(* Logix 5000 project; controller NWGG 1756-L72 rev 35.12; software revision 35.00 *)

TASK _2_MAIN (event, rate 10 ms, priority 15, watchdog 500 ms) : _2_MAIN
TASK Development (event, rate 10 ms, priority 10, watchdog 500 ms) : Main
TASK MainTask (continuous, watchdog 500 ms) : MainProgram
TASK SeedCleaning (event, rate 10 ms, priority 10, watchdog 500 ms) : Amp_Guages
TASK SeedLoadout (event, rate 10 ms, priority 10, watchdog 500 ms) : SeedLoadoutMain, Scale
TASK Test (event, rate 10 ms, priority 10, watchdog 500 ms) : Test
TASK UpdateBinConfig (event, rate 10 ms, priority 10, watchdog 500 ms)

MODULES
   Local : 1756-L72 (ICP 3, rev 35.12)
      R0S3_IA16 : 1756-IA16 (ICP 0, rev 3.1, Input RPI 20 ms)
      R0S2_IA16 : 1756-IA16 (ICP 1, rev 3.1, Input RPI 20 ms)
      R0S5_OA16I : 1756-OA16I (ICP 5, rev 3.1, Output RPI 20 ms)
      R0S6_OA16I : 1756-OA16I (ICP 6, rev 3.1, Output RPI 20 ms)
      R0S1_EN2TR : vendor 1 type 12 code 200 (ICP 4, Ethernet 192.10.21.33, rev 5.1)
         Treater_PLC : vendor 1 type 14 code 107 (Ethernet 192.10.21.15, rev 28.12, $43c9857a$ RPI 20 ms)
         LCP101_ETAP : 1783-ETAP (Ethernet 192.10.21.22, rev 2.1)
         Concrete_PLC : 1769-L35E Ethernet Port (Ethernet 192.10.21.32, rev 18.1)
            Concrete_PLC_Controller : vendor 1 type 14 code 65 (CompactLogixL35Controller 0, rev 18.1, $0a5c8464$ RPI 20 ms, $a6a510d7$ RPI 20 ms, $5be82f5e$ RPI 20 ms, $3e907429$ RPI 20 ms, $784e80a8$ RPI 20 ms, $ecd2168b$ RPI 100 ms, $00c6bec2$ RPI 20 ms, $fbd2347d$ RPI 20 ms, $adf8042c$ RPI 20 ms)
         Cimbria_Fan : PowerFlex 525-EENET (Ethernet 192.10.21.43, rev 4.1, Output RPI 20 ms)
         LCP103_4 : 1794-AENTR (Ethernet 192.10.21.39, rev 1.1, Output RPI 20 ms)
             : 1794-IA16 (Flex 2, rev 1.1)
            INPUT3 : 1794-IB16 (Flex 3, rev 1.1)
            CT_INPUT : 1794-IE12 (Flex 0, rev 1.1, Output RPI 80 ms)
            CT_INPUT2 : 1794-IE12 (Flex 1, rev 1.1, Output RPI 80 ms)
         R5M4_AENTR : 1794-AENTR (Ethernet 192.10.21.25, rev 1.1, Output RPI 20 ms)
            R5S3_IE8 : vendor 1 type 10 code 25 (Flex 3, rev 2.1, Input RPI 80 ms)
            R5S1_OE4 : 1794-OE4 (Flex 1, rev 2.1, Output RPI 80 ms)
            R5S0_OE4 : 1794-OE4 (Flex 0, rev 2.1, Output RPI 80 ms)
            R5S2_IE8 : vendor 1 type 10 code 25 (Flex 2, rev 2.1, Input RPI 80 ms)
         R4M2_AENTR : 1794-AENTR (Ethernet 192.10.21.27, rev 1.1, Output RPI 20 ms)
            R4S3_IA16 : 1794-IA16 (Flex 3, rev 1.1)
            R4S4_IA16 : 1794-IA16 (Flex 4, rev 1.1)
            R4SO_IA16 : 1794-IA16 (Flex 0, rev 1.1)
            R4S2_IA16 : 1794-IA16 (Flex 2, rev 1.1)
            R4S1_IA16 : 1794-IA16 (Flex 1, rev 1.1)
         DISTRIBUTION : 1794-AENTR (Ethernet 192.10.21.28, rev 1.1, Output RPI 20 ms)
            R5S1_OW8 : 1794-OW8 (Flex 1, rev 1.1)
            R5S0 : 1794-IA16 (Flex 0, rev 1.1)
         R4M3_AENTR : 1794-AENTR (Ethernet 192.10.21.26, rev 1.1, Output RPI 20 ms)
            R4S1_OA16 : vendor 1 type 7 code 48 (Flex 1, rev 1.1)
            R4S4_OA16 : vendor 1 type 7 code 48 (Flex 4, rev 1.1)
            R4S0_OA16 : vendor 1 type 7 code 48 (Flex 0, rev 1.1)
            R4S2_OA16 : vendor 1 type 7 code 48 (Flex 2, rev 1.1)
            R4S3_OA16 : vendor 1 type 7 code 48 (Flex 3, rev 1.1)
         R3M1_AENTR : 1794-AENTR (Ethernet 192.10.21.24, rev 1.1, Output RPI 20 ms)
            R3S1_OA16 : vendor 1 type 7 code 48 (Flex 1, rev 1.1)
            R3S3_OA16 : vendor 1 type 7 code 48 (Flex 3, rev 1.1)
            R3S0_IA16 : 1794-IA16 (Flex 0, rev 1.1)
            R3S2_IA16 : 1794-IA16 (Flex 2, rev 1.1)
         Stratix_5700 : vendor 1 type 12 code 241 (Ethernet 192.10.21.200, rev 4.1, Output RPI 1000 ms)
         AveryWT_Bay1 : ETHERNET-MODULE (Ethernet 192.10.21.70, rev 1.1, Output RPI 10 ms)
         AveryWT_Bay2 : ETHERNET-MODULE (Ethernet 192.10.21.71, rev 1.1, Output RPI 10 ms)
         R2S0_AENTR : vendor 1 type 12 code 228 (Ethernet 192.10.21.21, rev 1.1)
            R2S3_NI8 : vendor 1 type 117 code 6 (SLCChassis 3, rev 1.1, StandardDataDriven RPI 20 ms)
            R2S1_OA16 : vendor 1 type 116 code 24 (SLCChassis 1, rev 1.1, StandardDataDriven RPI 20 ms)
            R2S4_NI8 : vendor 1 type 117 code 6 (SLCChassis 4, rev 1.1, StandardDataDriven RPI 20 ms)
            R2S5_NI8 : vendor 1 type 117 code 6 (SLCChassis 5, rev 1.1, StandardDataDriven RPI 20 ms)
         R1S0_AENTR : vendor 1 type 12 code 228 (Ethernet 192.10.21.20, rev 1.1)
            R1S5_IA16 : vendor 1 type 116 code 3 (SLCChassis 5, rev 1.1, StandardDataDriven RPI 20 ms)
            R1S9_OA161 : vendor 1 type 116 code 24 (SLCChassis 10, rev 1.1, StandardDataDriven RPI 20 ms)
            R1S2_IA16 : vendor 1 type 116 code 3 (SLCChassis 2, rev 1.1, StandardDataDriven RPI 20 ms)
            R1S6_IA16 : vendor 1 type 116 code 3 (SLCChassis 6, rev 1.1, StandardDataDriven RPI 20 ms)
            R1S4_IA16 : vendor 1 type 116 code 3 (SLCChassis 4, rev 1.1, StandardDataDriven RPI 20 ms)
            R1S7_IA16 : vendor 1 type 116 code 3 (SLCChassis 7, rev 1.1, StandardDataDriven RPI 20 ms)
            R1S9_OA163 : vendor 1 type 116 code 24 (SLCChassis 12, rev 1.1, StandardDataDriven RPI 20 ms)
            R1S1_IA16 : vendor 1 type 116 code 3 (SLCChassis 1, rev 1.1, StandardDataDriven RPI 20 ms)
            R1S8_IA16 : vendor 1 type 116 code 3 (SLCChassis 8, rev 1.1, StandardDataDriven RPI 20 ms)
            R1S9_OA162 : vendor 1 type 116 code 24 (SLCChassis 11, rev 1.1, StandardDataDriven RPI 20 ms)
            R1S9_OA16 : vendor 1 type 116 code 24 (SLCChassis 9, rev 1.1, StandardDataDriven RPI 20 ms)
            R1S3_IA16 : vendor 1 type 116 code 3 (SLCChassis 3, rev 1.1, StandardDataDriven RPI 20 ms)
      Analog_Input : 1756-IF8 (ICP 2, rev 1.1, Input RPI 100 ms)
END_MODULES

TYPE udt_Andco_Remote_Out :
STRUCT
   Close : BOOL;
   Open : BOOL;
END_STRUCT
END_TYPE

TYPE udt_Andco_Values :
STRUCT
   Faulted : BOOL;
   Closed : BOOL;
   Values_Updated : BOOL;
   Fully_Open : BOOL;
   Com_Fault : BOOL;
   Open_Gate : BOOL;
   Close_Gate : BOOL;
   Cal_Gate : BOOL;
   Move_Gate : BOOL;
   Cal_Status : DINT;
   Raw_Position : DINT;
   Max_Position : DINT;
   Preact : DINT;
   Tolerance : DINT;
   Percent_Open : REAL;
   New_Pos : INT;
   Width : REAL;
   Rate : REAL;
   Pounds_Per_Inch : REAL;
   New_Rate : REAL;
   Set_New_Rate : BOOL;
   Display_New_Rate_Screen : BOOL;
   Analog : BOOL;
   Min_Position : DINT;
   Length : REAL;
   InchesOpen : REAL;
   AnalogValue : DINT;
END_STRUCT
END_TYPE

TYPE udt_Bin_Rate_Cal_Points :
STRUCT
   Andco_Position : INT;
   Rate : INT;
END_STRUCT
END_TYPE

TYPE udt_Clean_Seed_Bin :
STRUCT
   In_Use : BOOL;
   Bin_Name : STRING;
   Andco : udt_Andco_Values;
   Required_Clean_Belt : DINT;
   Required_Treat_Belt : DINT;
   Required_Transfer_Belt : DINT;
   Clean_Legs_Rqd : DINT;
   K_Valves_On_Treat : DINT;
   K_Valves_On_Clean : DINT;
   Concrete_Bin : BOOL;
   High_Bindicator : BOOL;
   Low_Bindicator : BOOL;
   Use_For_Clean : BOOL;
   Use_For_Treated : BOOL;
   Use_For_Transfer : BOOL;
   Cal_Mode : BOOL;
   Time_To_Treater : REAL;
   Time_To_Clean : REAL;
   Auger : BOOL;
   Current_Product : STRING;
   Capacity : DINT;
   Current_Amount : DINT;
END_STRUCT
END_TYPE

TYPE udt_Color :
STRUCT
   Color : INT;
   Duration : INT;
END_STRUCT
END_TYPE

TYPE udt_Cyclone :
STRUCT
   Start_Both_Fans : BOOL;
   Start_Cyclone : BOOL;
   Start_Aspirator : BOOL;
   Both_Fans_Running : BOOL;
   Cyclone_Running : BOOL;
   Aspirator_Running : BOOL;
END_STRUCT
END_TYPE

TYPE udt_Loadout_Air_Gate_Open :
STRUCT
   Manual_Open : BOOL;
   Auto_Open : BOOL;
   Auto_Open_Request : BOOL;
END_STRUCT
END_TYPE

TYPE udt_Loadout_Bin :
STRUCT
   Bin_Description : STRING;
   Bin_Variety : Variety;
   Manual_Open : BOOL;
   Air_Gate_Opened : BOOL;
   Use_For_Clean_Loadout : BOOL;
   Use_For_Treat_Loadout : BOOL;
   Use_For_Transfer_To : BOOL;
   Cal_Bin : BOOL;
   Rate_Cal_Points : udt_Bin_Rate_Cal_Points[6];
   InActive : BOOL;
   Clean_Load_Delay_Start : DINT;
   Treat_Load_Delay_Start : DINT;
   Bindicator_Low : BOOL;
   Air_Gate_Opening : BOOL;
   Andco_Values : udt_Andco_Values;
   Clean_Load_Delay_Stop : DINT;
   Treat_Load_Delay_Stop : DINT;
   Use_For_Transfer_From : BOOL;
   Can_Use_For_Transfer : BOOL;
   Selectable : BOOL;
   Temp_Rate_Cal_Points : udt_Bin_Rate_Cal_Points[6];
   Treat_Load_Delay : BOOL;
   tmrStartDelay : TIMER;
   tmrStopDelay : TIMER;
   StartDelayPre : INT;
   StopDelayPre : INT;
   Available_For_Clean_Load : BOOL;
   Available_For_Treat_Load : BOOL;
END_STRUCT
END_TYPE

TYPE udt_Loadout_K_Valve :
STRUCT
   Send_To_Treater : BOOL;
   Treater_Gate_Opened : BOOL;
   Clean_Gate_Opened : BOOL;
   One_Relay_Only : BOOL;
   Status_State : INT;
   Gate_Moving : BOOL;
END_STRUCT
END_TYPE

TYPE udt_Motor :
STRUCT
   Motor_Start : udt_Motor_Start;
   Motor_Control : Motor_Control;
   Running : BOOL;
   Motor_Config : udt_Motor_Config;
   Starting : BOOL;
   Run_Mode : DINT;
   Request_Auto_Start : BOOL;
END_STRUCT
END_TYPE

TYPE udt_Motor_Config :
STRUCT
   Definition : STRING;
   Wind_Up_Time : DINT;
   Stop_When_Plugged : BOOL;
   Stop_At_SLP20 : BOOL;
   Stop_At_Max_Amps : BOOL;
   Max_Amps : REAL;
   Speed_Sensor_Disabled : BOOL;
   Plugged_Sensor_Disabled : BOOL;
   Min_Motor_Amps : REAL;
   Warning_Amps : REAL;
END_STRUCT
END_TYPE

TYPE udt_Motor_Remote_In :
STRUCT
   Spd_20_Out : BOOL;
   Spd_10_Out : BOOL;
   Amps : REAL;
   Plug_Sensor : BOOL;
END_STRUCT
END_TYPE

TYPE udt_Motor_Start :
STRUCT
   Start_Motor : BOOL;
   Delay_Start : BOOL;
   Auto_Stop_Delay : INT;
   Required_For_Clean_Batch : BOOL;
   Required_For_Treat_Batch : BOOL;
   Required_For_Transfer_Batch : BOOL;
   Required_For_Cal : BOOL;
END_STRUCT
END_TYPE

TYPE udt_Not_Used :
STRUCT
   Always_ON : BOOL;
   Always_Off : BOOL;
   Always_Zero : DINT;
END_STRUCT
END_TYPE

TYPE udt_Requested_Variety :
STRUCT
   Item_Number : STRING;
   Percentage : REAL;
   Bin_Available : BOOL;
   In_Use : BOOL;
END_STRUCT
END_TYPE

TYPE udt_Treater_Loadout :
STRUCT
   Use_A_Treater : BOOL;
   Use_B_Treater : BOOL;
   Treater_Loadout_State : INT;
   Treater_Rate : INT;
   Auto_Start : BOOL;
   Manual_Start : BOOL;
   Close_Drip_Gate_Manual : BOOL;
   Drip_Gate_Closed : BOOL;
END_STRUCT
END_TYPE

TYPE udt_Truck_Scale :
STRUCT
   Description : STRING;
   Gross : REAL;
   Rate : REAL;
   Rate_Stable : BOOL;
   Avg_Rate : REAL;
   Rate_Tol : REAL;
   Error_Code : INT;
   Faulted : BOOL;
   Int_Rate : INT;
END_STRUCT
END_TYPE

TYPE Varieties_DB :
STRUCT
   Id : DINT;
   Name : STRING;
   ClassId : DINT;
   ClassType : STRING;
   MarketClassId : DINT;
   MarketClassType : STRING;
   Breeder : STRING;
   Trate : STRING;
   FullDecription : STRING;
END_STRUCT
END_TYPE

TYPE Variety :
STRUCT
   Item_Number : STRING;
   Name : STRING;
   Class : STRING;
   Color : udt_Color[4];
END_STRUCT
END_TYPE

ADD_ON_INSTRUCTION AI   (* revision 1.0, vendor Rockwell Automation *)
VAR_INPUT
   In : ALIAS FOR SCL_01.In; {access None, required}
   RawMin : ALIAS FOR SCL_01.InRawMin; {access None, required}
   RawMax : ALIAS FOR SCL_01.InRawMax; {access None, required}
   EUMin : ALIAS FOR SCL_01.InEUMin; {access None, required}
   EUMax : ALIAS FOR SCL_01.InEUMax; {access None, required}
END_VAR
VAR_OUTPUT
   Out : ALIAS FOR SCL_01.Out; {access None, required}
END_VAR
VAR
   SCL_01 : SCALE; {access None}
END_VAR

ROUTINE Logic   (* function block diagram *)
   SHEET 1
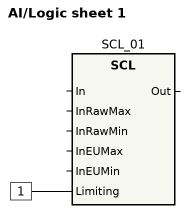
   SCL_01 : SCL(Limiting := 1);   // unwired pins: In InRawMax InRawMin InEUMax InEUMin Out
END_ROUTINE
END_ADD_ON_INSTRUCTION

ADD_ON_INSTRUCTION AI_SCALE   (* revision 1.0, vendor Rockwell Automation *)
VAR_INPUT
   In : ALIAS FOR SCL_01.In; {access None, required}
   RawMin : ALIAS FOR SCL_01.InRawMin; {access None, required}
   RawMax : ALIAS FOR SCL_01.InRawMax; {access None, required}
   EUMin : ALIAS FOR SCL_01.InEUMin; {access None, required}
   EUMax : ALIAS FOR SCL_01.InEUMax; {access None, required}
END_VAR
VAR_OUTPUT
   Out : ALIAS FOR SCL_01.Out; {access None, required}
END_VAR
VAR
   SCL_01 : SCALE; {access None}
END_VAR

ROUTINE Logic   (* function block diagram *)
   SHEET 1
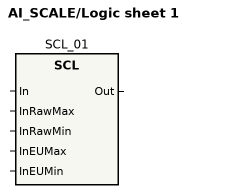
   SCL_01 : SCL();   // unwired pins: In InRawMax InRawMin InEUMax InEUMin Out
END_ROUTINE
END_ADD_ON_INSTRUCTION

ADD_ON_INSTRUCTION Andco   (* revision 1.0 *)
VAR_IN_OUT
   Andco_Values : udt_Andco_Values; {required}
   Andco_Motor_Open : BOOL; {required}
   Anco_Motor_Close : BOOL; {required}
END_VAR
VAR
   tmr_Web_Watchdog : TIMER := (PRE := 30000); {access None}
   Cal_Open_Gate : BOOL; {access None}
   Cal_Close_Gate : BOOL; {access None}
   ONS_Start_Calibration : BOOL; {access None}
   Motor_Wind_Down : DINT; {access None}
   Cal_Mid_Point : DINT; {access None}
   Cal_Preact : BOOL; {access None}
   Cal_Finish_Close_Gate : BOOL; {access None}
   tmr_Motor_Wind_Down : TIMER[8]; {access None}
   New_Position : DINT; {access None}
   Move_Open : BOOL; {access None}
   Move_Close : BOOL; {access None}
   Adjusted_New_Position : DINT; {access None}
   Cal_Init_Bin_Closed : BOOL; {access None}
END_VAR

ROUTINE Logic   (* ladder *)
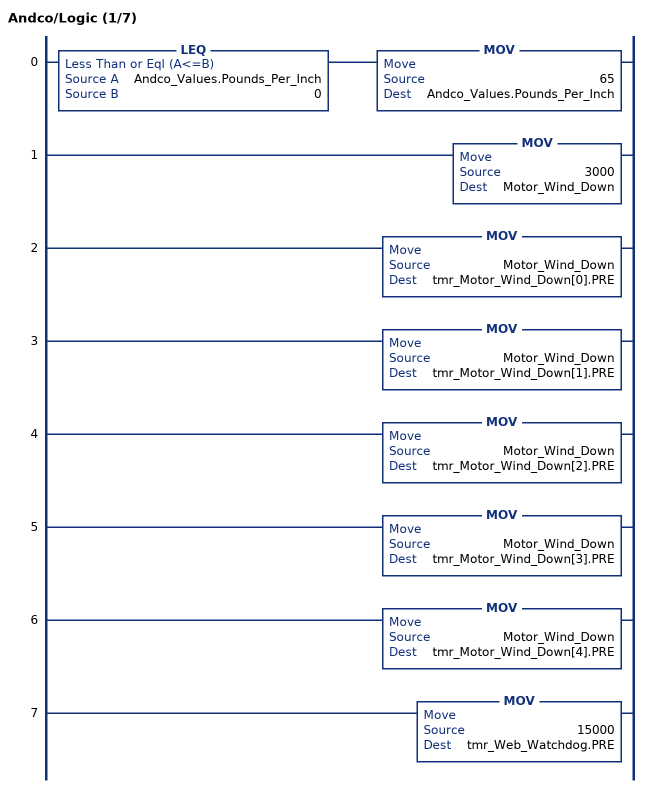
   0: LEQ(Andco_Values.Pounds_Per_Inch,0)MOV(65,Andco_Values.Pounds_Per_Inch);
   1: MOV(3000,Motor_Wind_Down);
   2: MOV(Motor_Wind_Down,tmr_Motor_Wind_Down[0].PRE);
   3: MOV(Motor_Wind_Down,tmr_Motor_Wind_Down[1].PRE);
   4: MOV(Motor_Wind_Down,tmr_Motor_Wind_Down[2].PRE);
   5: MOV(Motor_Wind_Down,tmr_Motor_Wind_Down[3].PRE);
   6: MOV(Motor_Wind_Down,tmr_Motor_Wind_Down[4].PRE);
   7: MOV(15000,tmr_Web_Watchdog.PRE);
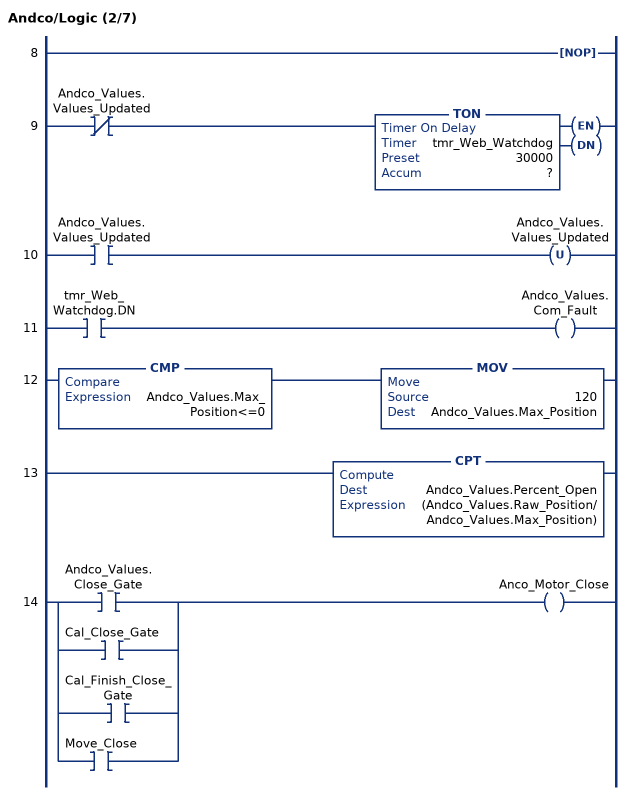
   8: NOP();
   9: XIO(Andco_Values.Values_Updated)TON(tmr_Web_Watchdog,?,?);
   10: XIC(Andco_Values.Values_Updated)OTU(Andco_Values.Values_Updated);
   11: XIC(tmr_Web_Watchdog.DN)OTE(Andco_Values.Com_Fault);
   12: CMP(Andco_Values.Max_Position<=0)MOV(120,Andco_Values.Max_Position);
   13: CPT(Andco_Values.Percent_Open,(Andco_Values.Raw_Position/Andco_Values.Max_Position));
   14: [XIC(Andco_Values.Close_Gate) ,XIC(Cal_Close_Gate) ,XIC(Cal_Finish_Close_Gate) ,XIC(Move_Close) ]OTE(Anco_Motor_Close);
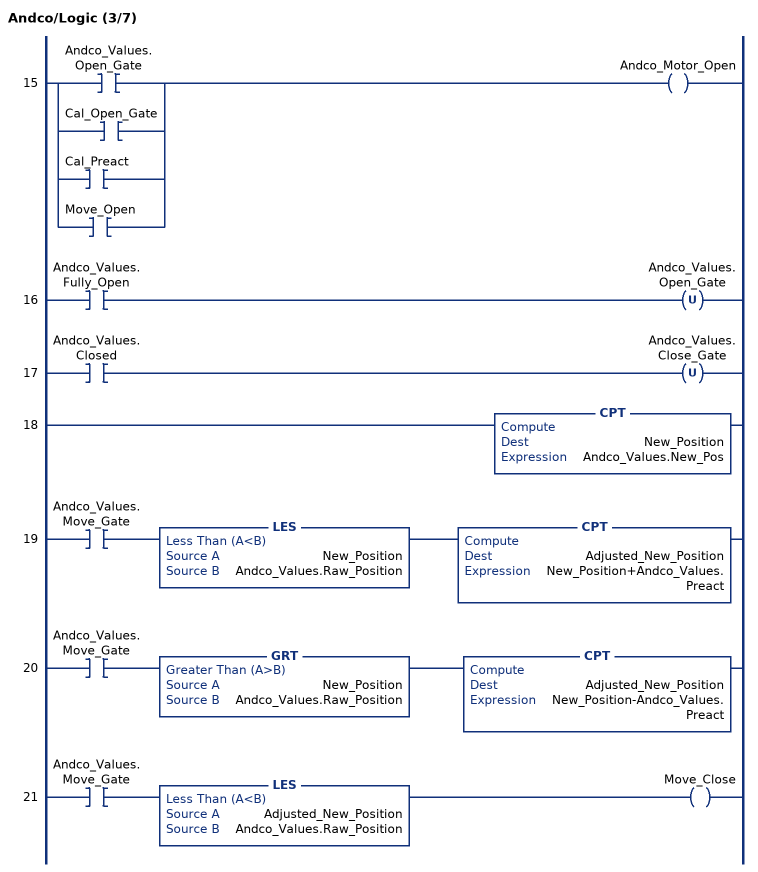
   15: [XIC(Andco_Values.Open_Gate) ,XIC(Cal_Open_Gate) ,XIC(Cal_Preact) ,XIC(Move_Open) ]OTE(Andco_Motor_Open);
   16: XIC(Andco_Values.Fully_Open)OTU(Andco_Values.Open_Gate);
   17: XIC(Andco_Values.Closed)OTU(Andco_Values.Close_Gate);
   18: CPT(New_Position,Andco_Values.New_Pos);
   19: XIC(Andco_Values.Move_Gate)LES(New_Position,Andco_Values.Raw_Position)CPT(Adjusted_New_Position,New_Position+Andco_Values.Preact);
   20: XIC(Andco_Values.Move_Gate)GRT(New_Position,Andco_Values.Raw_Position)CPT(Adjusted_New_Position,New_Position-Andco_Values.Preact);
   21: XIC(Andco_Values.Move_Gate)LES(Adjusted_New_Position,Andco_Values.Raw_Position)OTE(Move_Close);
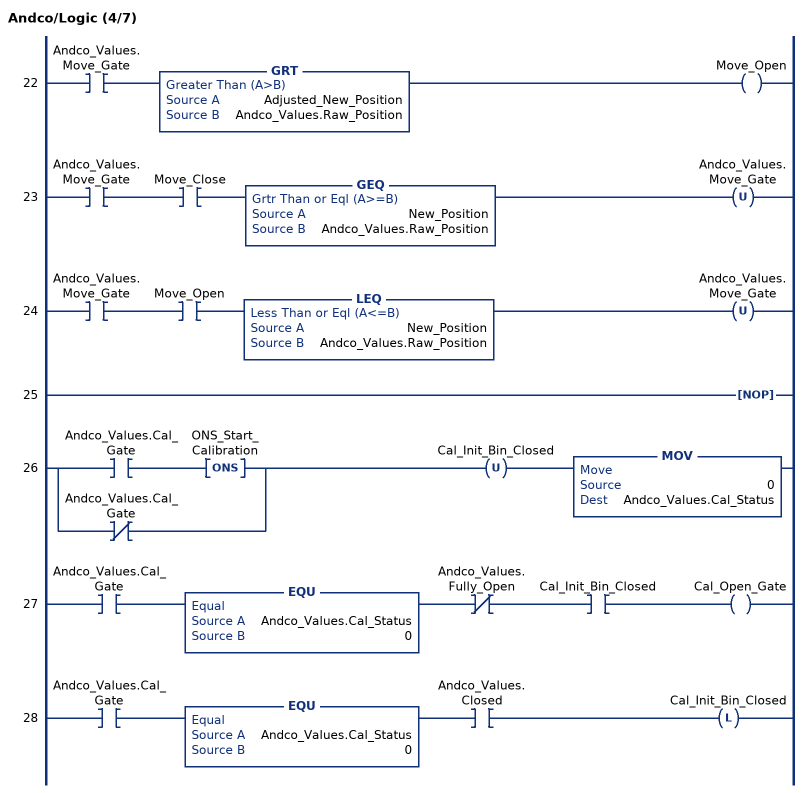
   22: XIC(Andco_Values.Move_Gate)GRT(Adjusted_New_Position,Andco_Values.Raw_Position)OTE(Move_Open);
   23: XIC(Andco_Values.Move_Gate)XIC(Move_Close)GEQ(New_Position,Andco_Values.Raw_Position)OTU(Andco_Values.Move_Gate);
   24: XIC(Andco_Values.Move_Gate)XIC(Move_Open)LEQ(New_Position,Andco_Values.Raw_Position)OTU(Andco_Values.Move_Gate);
   25: NOP();
   26: [XIC(Andco_Values.Cal_Gate) ONS(ONS_Start_Calibration) ,XIO(Andco_Values.Cal_Gate) ]OTU(Cal_Init_Bin_Closed)MOV(0,Andco_Values.Cal_Status);
   27: XIC(Andco_Values.Cal_Gate)EQU(Andco_Values.Cal_Status,0)XIO(Andco_Values.Fully_Open)XIC(Cal_Init_Bin_Closed)OTE(Cal_Open_Gate);
   28: XIC(Andco_Values.Cal_Gate)EQU(Andco_Values.Cal_Status,0)XIC(Andco_Values.Closed)OTL(Cal_Init_Bin_Closed);
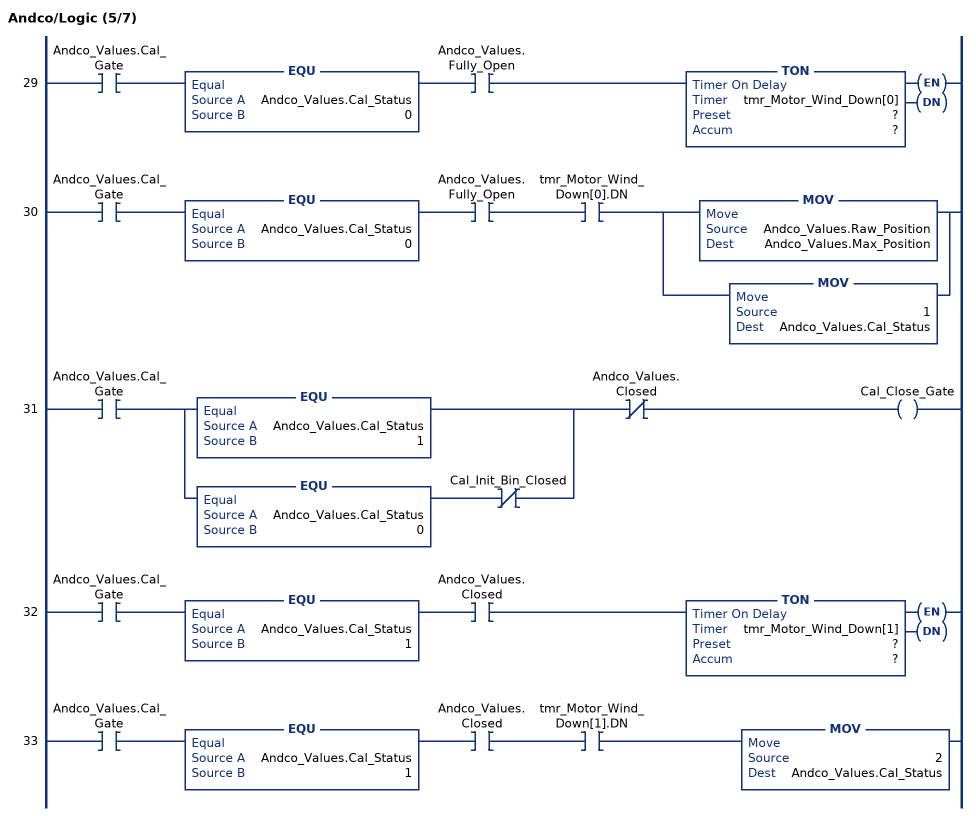
   29: XIC(Andco_Values.Cal_Gate)EQU(Andco_Values.Cal_Status,0)XIC(Andco_Values.Fully_Open)TON(tmr_Motor_Wind_Down[0],?,?);
   30: XIC(Andco_Values.Cal_Gate)EQU(Andco_Values.Cal_Status,0)XIC(Andco_Values.Fully_Open)XIC(tmr_Motor_Wind_Down[0].DN)[MOV(Andco_Values.Raw_Position,Andco_Values.Max_Position) ,MOV(1,Andco_Values.Cal_Status) ];
   31: XIC(Andco_Values.Cal_Gate)[EQU(Andco_Values.Cal_Status,1) ,EQU(Andco_Values.Cal_Status,0) XIO(Cal_Init_Bin_Closed) ]XIO(Andco_Values.Closed)OTE(Cal_Close_Gate);
   32: XIC(Andco_Values.Cal_Gate)EQU(Andco_Values.Cal_Status,1)XIC(Andco_Values.Closed)TON(tmr_Motor_Wind_Down[1],?,?);
   33: XIC(Andco_Values.Cal_Gate)EQU(Andco_Values.Cal_Status,1)XIC(Andco_Values.Closed)XIC(tmr_Motor_Wind_Down[1].DN)MOV(2,Andco_Values.Cal_Status);
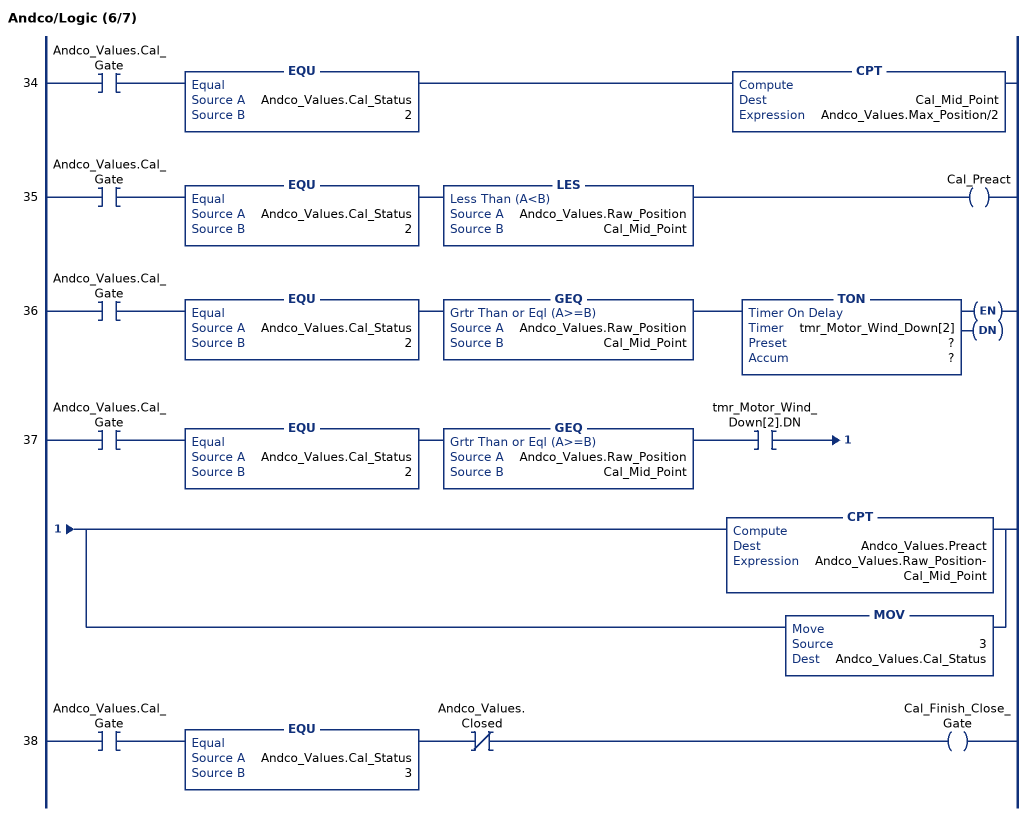
   34: XIC(Andco_Values.Cal_Gate)EQU(Andco_Values.Cal_Status,2)CPT(Cal_Mid_Point,Andco_Values.Max_Position/2);
   35: XIC(Andco_Values.Cal_Gate)EQU(Andco_Values.Cal_Status,2)LES(Andco_Values.Raw_Position,Cal_Mid_Point)OTE(Cal_Preact);
   36: XIC(Andco_Values.Cal_Gate)EQU(Andco_Values.Cal_Status,2)GEQ(Andco_Values.Raw_Position,Cal_Mid_Point)TON(tmr_Motor_Wind_Down[2],?,?);
   37: XIC(Andco_Values.Cal_Gate)EQU(Andco_Values.Cal_Status,2)GEQ(Andco_Values.Raw_Position,Cal_Mid_Point)XIC(tmr_Motor_Wind_Down[2].DN)[CPT(Andco_Values.Preact,Andco_Values.Raw_Position-Cal_Mid_Point) ,MOV(3,Andco_Values.Cal_Status) ];
   38: XIC(Andco_Values.Cal_Gate)EQU(Andco_Values.Cal_Status,3)XIO(Andco_Values.Closed)OTE(Cal_Finish_Close_Gate);
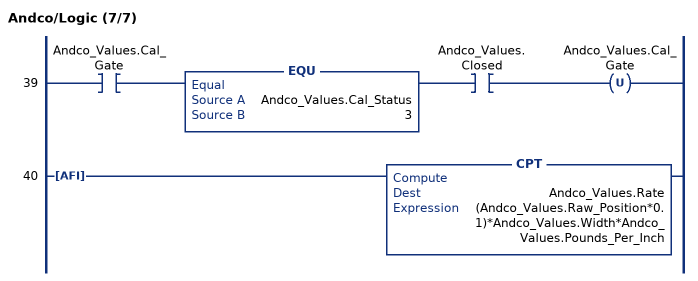
   39: XIC(Andco_Values.Cal_Gate)EQU(Andco_Values.Cal_Status,3)XIC(Andco_Values.Closed)OTU(Andco_Values.Cal_Gate);
   40: AFI()CPT(Andco_Values.Rate,(Andco_Values.Raw_Position*0.1)*Andco_Values.Width*Andco_Values.Pounds_Per_Inch);
END_ROUTINE
END_ADD_ON_INSTRUCTION

ADD_ON_INSTRUCTION AndcoAnalog   (* revision 1.0 *)
VAR_IN_OUT
   Andco_Values : udt_Andco_Values; {required}
   Andco_Motor_Open : BOOL; {required}
   Anco_Motor_Close : BOOL; {required}
END_VAR
VAR_INPUT
   AnalogValue : DINT; {access Read Only, required}
END_VAR
VAR
   tmr_Web_Watchdog : TIMER := (PRE := 30000); {access None}
   Cal_Open_Gate : BOOL; {access None}
   Cal_Close_Gate : BOOL; {access None}
   Motor_Wind_Down : DINT; {access None}
   Cal_Mid_Point : DINT; {access None}
   Cal_Preact : BOOL; {access None}
   Cal_Finish_Close_Gate : BOOL; {access None}
   tmr_Motor_Wind_Down : TIMER[8] := ([1].PRE := 1000, [2].PRE := 1000); {access None}
   New_Position : DINT; {access None}
   Move_Open : BOOL; {access None}
   Move_Close : BOOL; {access None}
   Adjusted_New_Position : DINT; {access None}
   Cal_Init_Bin_Closed : BOOL; {access None}
   tmrCalCloseGate : TIMER := (PRE := 55000); {access None}
   CurrentPosition : DINT; {access None}
   tmrCalOpenGate : TIMER := (PRE := 55000); {access None}
   CalReturnToPosition : BOOL; {access None}
   CalibratingGate : BOOL; {access None}
   onsStartCal : BOOL; {access None}
   sbCalGateClosed : BOOL; {access None}
   obCalGateClosed : BOOL; {access None}
   sbStartCal : BOOL; {access None}
   obStartCal : BOOL; {access None}
   sbCalGateOpened : BOOL; {access None}
   obCalGateOpened : BOOL; {access None}
END_VAR

ROUTINE Logic   (* ladder *)
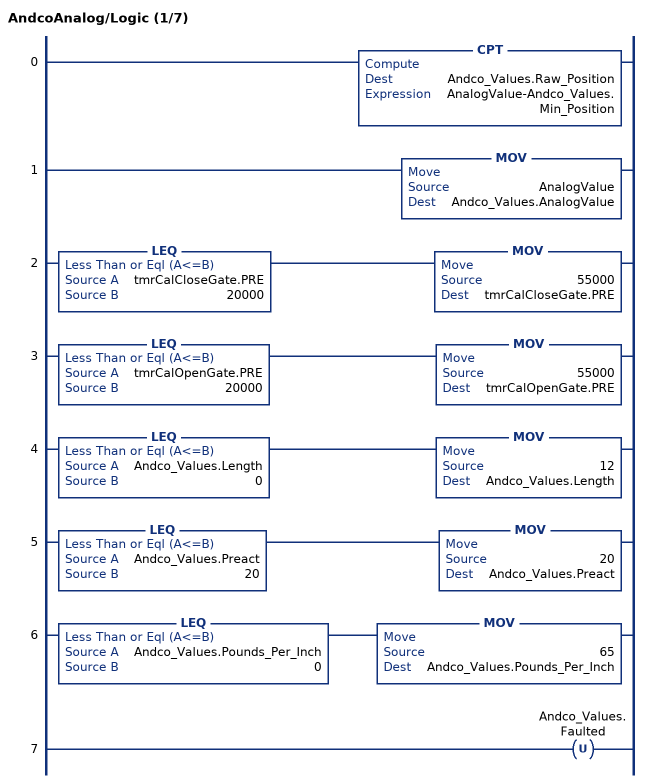
   0: CPT(Andco_Values.Raw_Position,AnalogValue-Andco_Values.Min_Position);
   1: MOV(AnalogValue,Andco_Values.AnalogValue);
   2: LEQ(tmrCalCloseGate.PRE,20000)MOV(55000,tmrCalCloseGate.PRE);
   3: LEQ(tmrCalOpenGate.PRE,20000)MOV(55000,tmrCalOpenGate.PRE);
   4: LEQ(Andco_Values.Length,0)MOV(12,Andco_Values.Length);
   5: LEQ(Andco_Values.Preact,20)MOV(20,Andco_Values.Preact);
   6: LEQ(Andco_Values.Pounds_Per_Inch,0)MOV(65,Andco_Values.Pounds_Per_Inch);
   7: OTU(Andco_Values.Faulted);
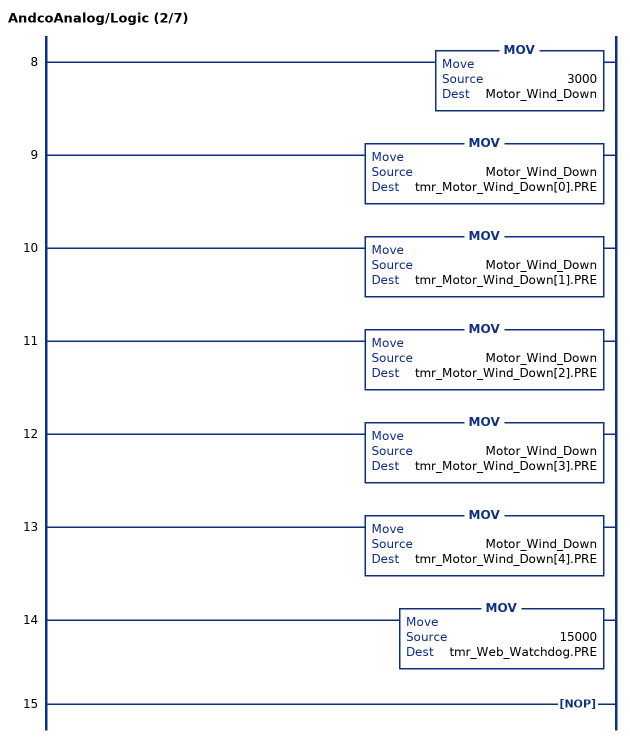
   8: MOV(3000,Motor_Wind_Down);
   9: MOV(Motor_Wind_Down,tmr_Motor_Wind_Down[0].PRE);
   10: MOV(Motor_Wind_Down,tmr_Motor_Wind_Down[1].PRE);
   11: MOV(Motor_Wind_Down,tmr_Motor_Wind_Down[2].PRE);
   12: MOV(Motor_Wind_Down,tmr_Motor_Wind_Down[3].PRE);
   13: MOV(Motor_Wind_Down,tmr_Motor_Wind_Down[4].PRE);
   14: MOV(15000,tmr_Web_Watchdog.PRE);
   15: NOP();
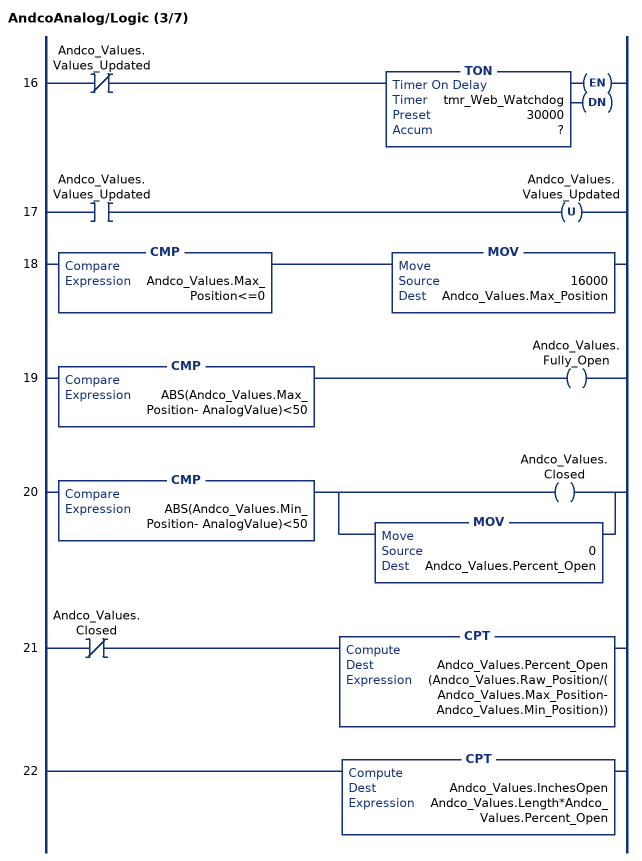
   16: XIO(Andco_Values.Values_Updated)TON(tmr_Web_Watchdog,?,?);
   17: XIC(Andco_Values.Values_Updated)OTU(Andco_Values.Values_Updated);
   18: CMP(Andco_Values.Max_Position<=0)MOV(16000,Andco_Values.Max_Position);
   19: CMP(ABS(Andco_Values.Max_Position- AnalogValue)<50)OTE(Andco_Values.Fully_Open);
   20: CMP(ABS(Andco_Values.Min_Position- AnalogValue)<50)[OTE(Andco_Values.Closed) ,MOV(0,Andco_Values.Percent_Open) ];
   21: XIO(Andco_Values.Closed)CPT(Andco_Values.Percent_Open,(Andco_Values.Raw_Position/(Andco_Values.Max_Position-Andco_Values.Min_Position)));
   22: CPT(Andco_Values.InchesOpen,Andco_Values.Length*Andco_Values.Percent_Open);
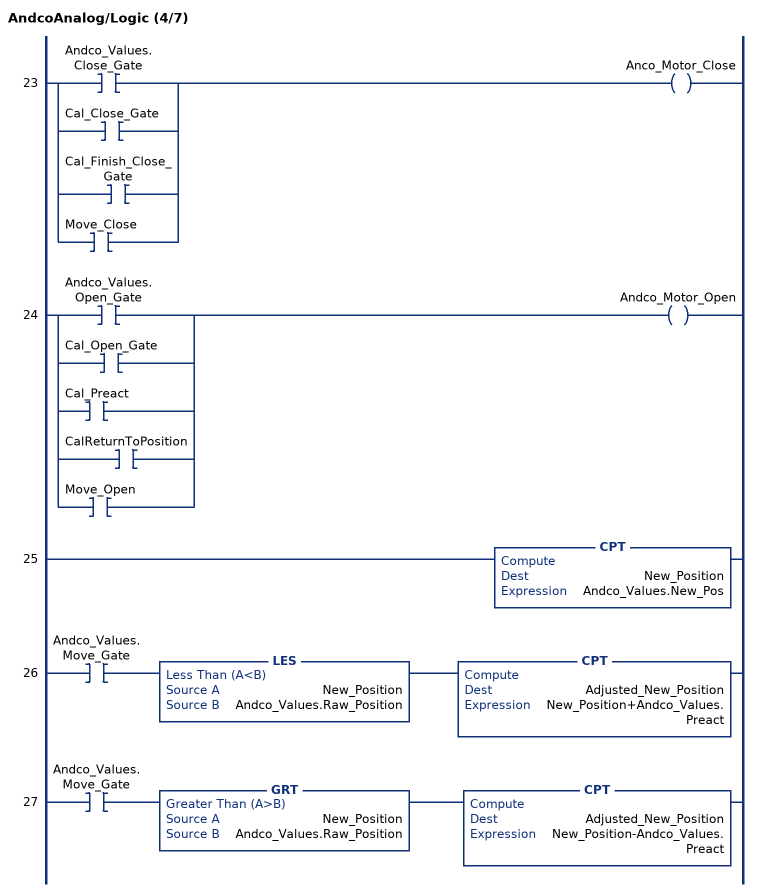
   23: [XIC(Andco_Values.Close_Gate) ,XIC(Cal_Close_Gate) ,XIC(Cal_Finish_Close_Gate) ,XIC(Move_Close) ]OTE(Anco_Motor_Close);
   24: [XIC(Andco_Values.Open_Gate) ,XIC(Cal_Open_Gate) ,XIC(Cal_Preact) ,XIC(CalReturnToPosition) ,XIC(Move_Open) ]OTE(Andco_Motor_Open);
   25: CPT(New_Position,Andco_Values.New_Pos);
   26: XIC(Andco_Values.Move_Gate)LES(New_Position,Andco_Values.Raw_Position)CPT(Adjusted_New_Position,New_Position+Andco_Values.Preact);
   27: XIC(Andco_Values.Move_Gate)GRT(New_Position,Andco_Values.Raw_Position)CPT(Adjusted_New_Position,New_Position-Andco_Values.Preact);
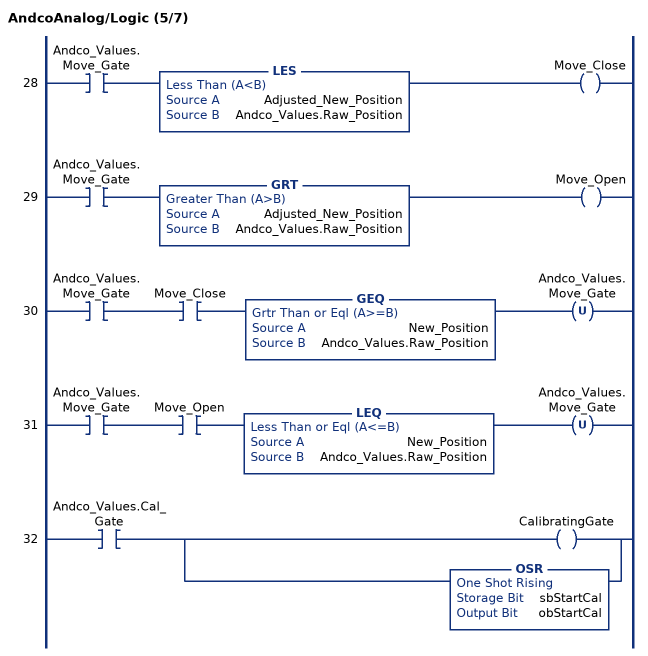
   28: XIC(Andco_Values.Move_Gate)LES(Adjusted_New_Position,Andco_Values.Raw_Position)OTE(Move_Close);
   29: XIC(Andco_Values.Move_Gate)GRT(Adjusted_New_Position,Andco_Values.Raw_Position)OTE(Move_Open);
   30: XIC(Andco_Values.Move_Gate)XIC(Move_Close)GEQ(New_Position,Andco_Values.Raw_Position)OTU(Andco_Values.Move_Gate);
   31: XIC(Andco_Values.Move_Gate)XIC(Move_Open)LEQ(New_Position,Andco_Values.Raw_Position)OTU(Andco_Values.Move_Gate);
   32: XIC(Andco_Values.Cal_Gate)[OTE(CalibratingGate) ,OSR(sbStartCal,obStartCal) ];
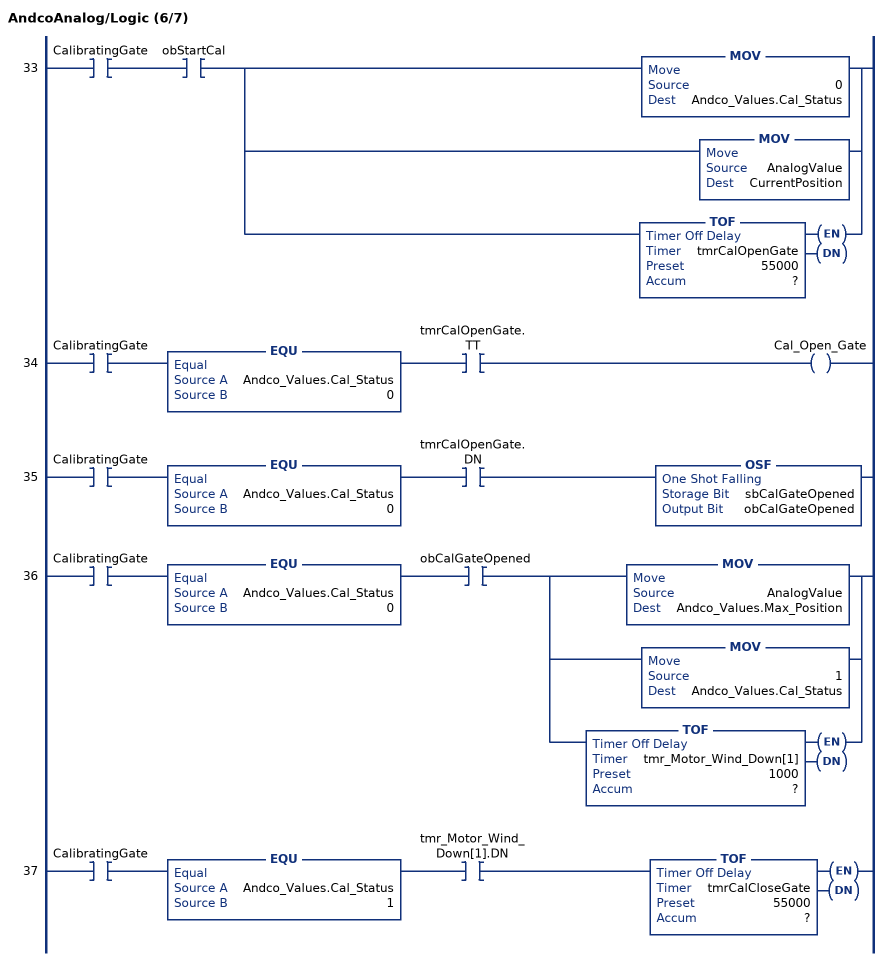
   33: XIC(CalibratingGate)XIC(obStartCal)[MOV(0,Andco_Values.Cal_Status) ,MOV(AnalogValue,CurrentPosition) ,TOF(tmrCalOpenGate,?,?) ];
   34: XIC(CalibratingGate)EQU(Andco_Values.Cal_Status,0)XIC(tmrCalOpenGate.TT)OTE(Cal_Open_Gate);
   35: XIC(CalibratingGate)EQU(Andco_Values.Cal_Status,0)XIC(tmrCalOpenGate.DN)OSF(sbCalGateOpened,obCalGateOpened);
   36: XIC(CalibratingGate)EQU(Andco_Values.Cal_Status,0)XIC(obCalGateOpened)[MOV(AnalogValue,Andco_Values.Max_Position) ,MOV(1,Andco_Values.Cal_Status) ,TOF(tmr_Motor_Wind_Down[1],?,?) ];
   37: XIC(CalibratingGate)EQU(Andco_Values.Cal_Status,1)XIC(tmr_Motor_Wind_Down[1].DN)TOF(tmrCalCloseGate,?,?);
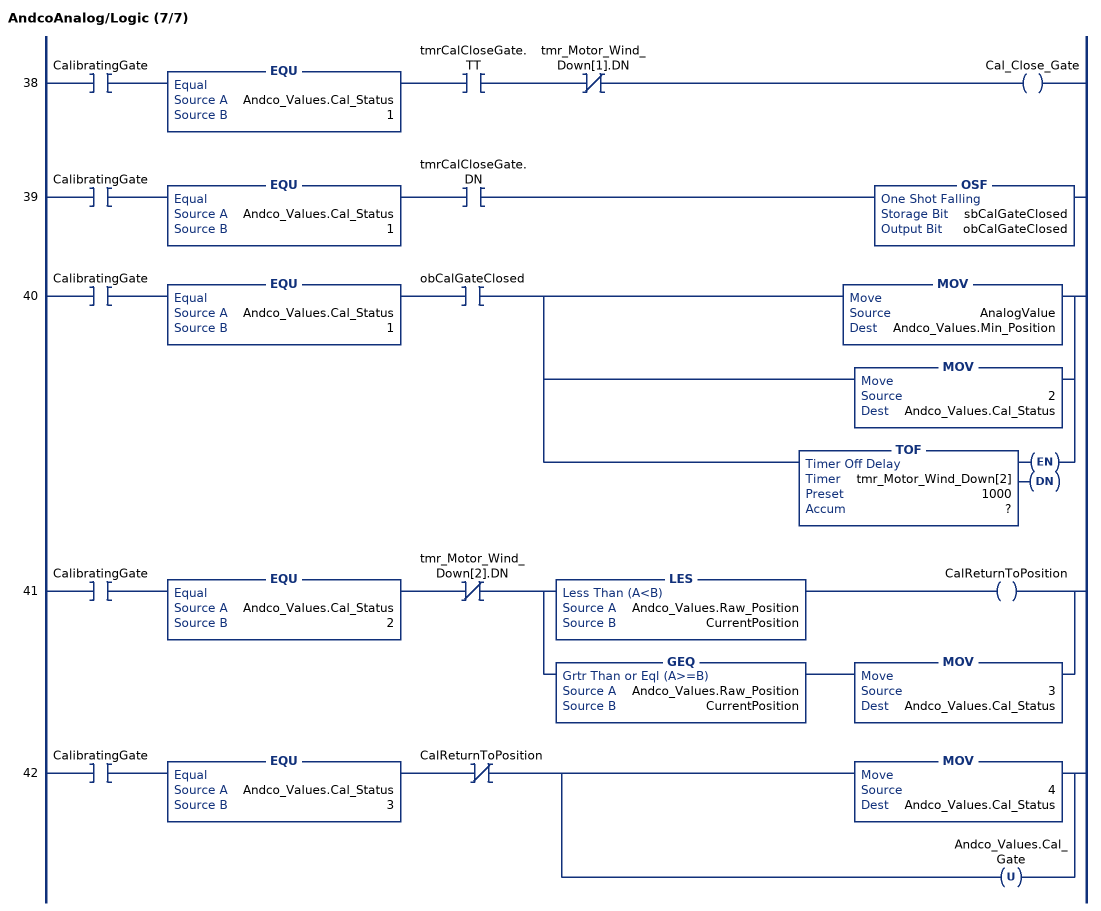
   38: XIC(CalibratingGate)EQU(Andco_Values.Cal_Status,1)XIC(tmrCalCloseGate.TT)XIO(tmr_Motor_Wind_Down[1].DN)OTE(Cal_Close_Gate);
   39: XIC(CalibratingGate)EQU(Andco_Values.Cal_Status,1)XIC(tmrCalCloseGate.DN)OSF(sbCalGateClosed,obCalGateClosed);
   40: XIC(CalibratingGate)EQU(Andco_Values.Cal_Status,1)XIC(obCalGateClosed)[MOV(AnalogValue,Andco_Values.Min_Position) ,MOV(2,Andco_Values.Cal_Status) ,TOF(tmr_Motor_Wind_Down[2],?,?) ];
   41: XIC(CalibratingGate)EQU(Andco_Values.Cal_Status,2)XIO(tmr_Motor_Wind_Down[2].DN)[LES(Andco_Values.Raw_Position,CurrentPosition) OTE(CalReturnToPosition) ,GEQ(Andco_Values.Raw_Position,CurrentPosition) MOV(3,Andco_Values.Cal_Status) ];
   42: XIC(CalibratingGate)EQU(Andco_Values.Cal_Status,3)XIO(CalReturnToPosition)[MOV(4,Andco_Values.Cal_Status) ,OTU(Andco_Values.Cal_Gate) ];
END_ROUTINE
END_ADD_ON_INSTRUCTION

ADD_ON_INSTRUCTION HOUR_METER   (* revision 1.0 *)
VAR_INPUT
   MOTOR_RUNNING_INPUT_1 : BOOL; {required}
END_VAR
VAR_OUTPUT
   HR_METER_DISPLAY : DINT; {visible}
END_VAR
VAR_INPUT
   NEXT_SCHDL_MAINTENANCE : DINT; {visible}
END_VAR
VAR_OUTPUT
   MAINTENANCE_ALARM : BOOL; {visible}
END_VAR
VAR
   COUNTER : COUNTER := (PRE := 99999999); {access None}
   TIMER : TIMER := (PRE := 3600000); {access None}
END_VAR

ROUTINE Logic   (* ladder *)
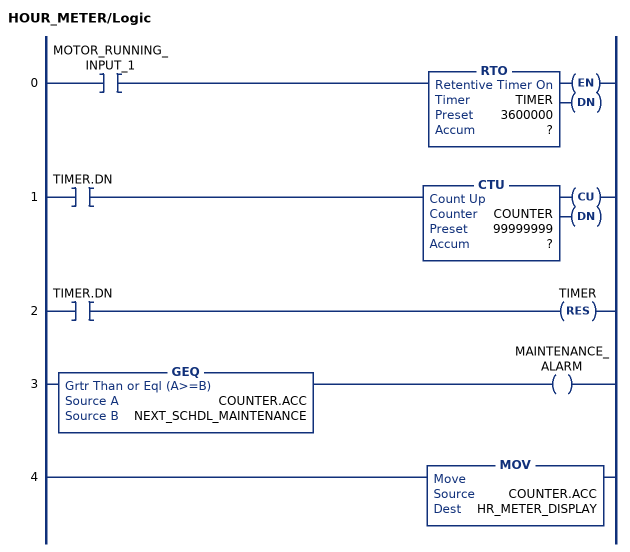
   0: XIC(MOTOR_RUNNING_INPUT_1)RTO(TIMER,?,?);
   1: XIC(TIMER.DN)CTU(COUNTER,?,?);
   2: XIC(TIMER.DN)RES(TIMER);
   3: GEQ(COUNTER.ACC,NEXT_SCHDL_MAINTENANCE)OTE(MAINTENANCE_ALARM);
   4: MOV(COUNTER.ACC,HR_METER_DISPLAY);
END_ROUTINE
END_ADD_ON_INSTRUCTION

ADD_ON_INSTRUCTION Loadout_Bin_Control   (* revision 1.0 *)
VAR_IN_OUT
   Bin : udt_Loadout_Bin; {required}
   Open_Air_Gate : BOOL; {required}
END_VAR
VAR_INPUT
   Bin_Open_Treat_Pause : BOOL; {required}
   Bin_Open_Clean_Pause : BOOL; {required}
END_VAR
VAR_IN_OUT
   TMR_Max_Treat_Delay : TIMER; {required}
   TMR_Max_Clean_Delay : TIMER; {required}
   Air_Gate_Open_Input : BOOL; {required}
   Auger_Relay : BOOL; {required}
END_VAR
VAR_INPUT
   Use_Auger_Relay : BOOL; {required}
   Use_Bindicator : BOOL; {access None, required}
END_VAR
VAR_IN_OUT
   Bindicator_Input : BOOL; {required}
   ALM_Air_Gate_Failed : ALARM_DIGITAL; {required}
END_VAR
VAR_INPUT
   Bin_Open_Transfer_Pause : BOOL; {required}
END_VAR
VAR_IN_OUT
   Clean_Batch_Status : DINT; {required}
   Treat_Batch_Status : DINT; {required}
   Transfer_Batch_Status : DINT; {required}
   Andco_Motor_Open : BOOL; {required}
   Andco_Motor_Close : BOOL; {required}
   Required_Belt : BOOL; {required}
   Manual_Mode : BOOL; {required}
END_VAR
VAR_INPUT
   RawAnalogTag : DINT; {access Read Only, required}
END_VAR
VAR
   Auto_Open_Air_Gate_Ready : BOOL; {access None}
   Air_Gate_Open_Cal : BOOL; {access None}
   TMR_Air_Gate_Fail : TIMER := (PRE := 4000); {access None}
   ALM_Air_Gate_Failed_Ack : BOOL; {access None}
   Air_Gate_Open_Clean : BOOL; {access None}
   Air_Gate_Open_Treat : BOOL; {access None}
   Air_Gate_Open_Transfer : BOOL; {access None}
   Andco : Andco; {access None}
   Open_Treat_Air_Gate : BOOL; {access None}
   Open_Treat_Air_Gate_Ready : BOOL; {access None}
   AndcoAnalog : AndcoAnalog; {access None}
END_VAR

ROUTINE Logic   (* ladder *)
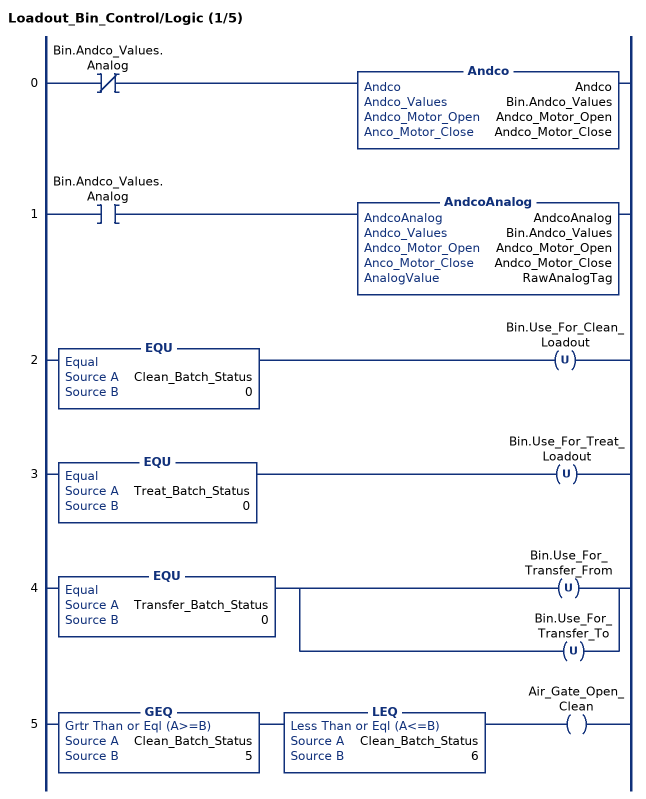
   0: XIO(Bin.Andco_Values.Analog)Andco(Andco,Bin.Andco_Values,Andco_Motor_Open,Andco_Motor_Close);
   1: XIC(Bin.Andco_Values.Analog)AndcoAnalog(AndcoAnalog,Bin.Andco_Values,Andco_Motor_Open,Andco_Motor_Close,RawAnalogTag);
   2: EQU(Clean_Batch_Status,0)OTU(Bin.Use_For_Clean_Loadout);
   3: EQU(Treat_Batch_Status,0)OTU(Bin.Use_For_Treat_Loadout);
   4: EQU(Transfer_Batch_Status,0)[OTU(Bin.Use_For_Transfer_From) ,OTU(Bin.Use_For_Transfer_To) ];
   5: GEQ(Clean_Batch_Status,5)LEQ(Clean_Batch_Status,6)OTE(Air_Gate_Open_Clean);
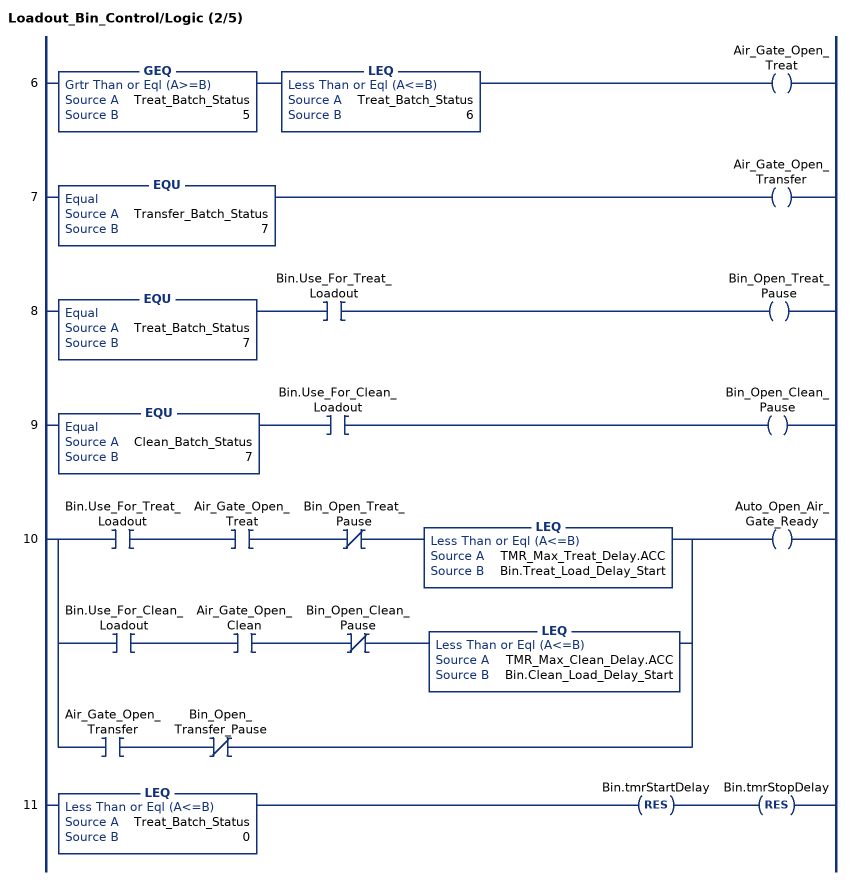
   6: GEQ(Treat_Batch_Status,5)LEQ(Treat_Batch_Status,6)OTE(Air_Gate_Open_Treat);
   7: EQU(Transfer_Batch_Status,7)OTE(Air_Gate_Open_Transfer);
   8: EQU(Treat_Batch_Status,7)XIC(Bin.Use_For_Treat_Loadout)OTE(Bin_Open_Treat_Pause);
   9: EQU(Clean_Batch_Status,7)XIC(Bin.Use_For_Clean_Loadout)OTE(Bin_Open_Clean_Pause);
   10: [XIC(Bin.Use_For_Treat_Loadout) XIC(Air_Gate_Open_Treat) XIO(Bin_Open_Treat_Pause) LEQ(TMR_Max_Treat_Delay.ACC,Bin.Treat_Load_Delay_Start) ,XIC(Bin.Use_For_Clean_Loadout) XIC(Air_Gate_Open_Clean) XIO(Bin_Open_Clean_Pause) LEQ(TMR_Max_Clean_Delay.ACC,Bin.Clean_Load_Delay_Start) ,XIC(Air_Gate_Open_Transfer) XIO(Bin_Open_Transfer_Pause) ]OTE(Auto_Open_Air_Gate_Ready);
   11: LEQ(Treat_Batch_Status,0)RES(Bin.tmrStartDelay)RES(Bin.tmrStopDelay);
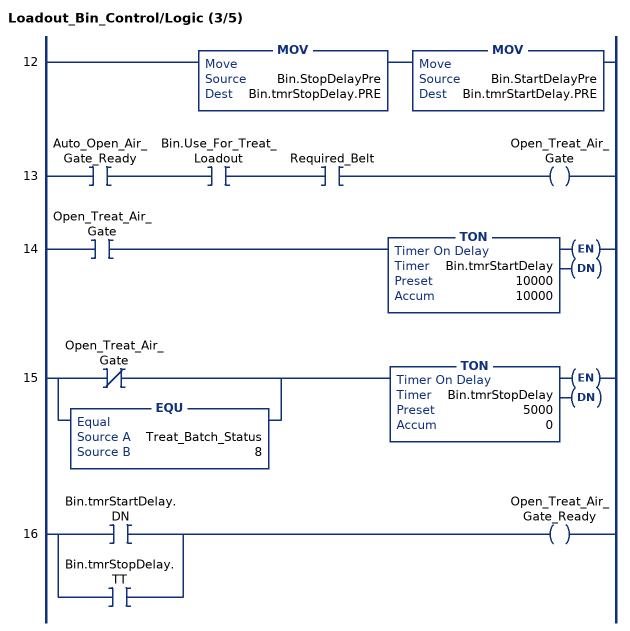
   12: MOV(Bin.StopDelayPre,Bin.tmrStopDelay.PRE)MOV(Bin.StartDelayPre,Bin.tmrStartDelay.PRE);
   13: XIC(Auto_Open_Air_Gate_Ready)XIC(Bin.Use_For_Treat_Loadout)XIC(Required_Belt)OTE(Open_Treat_Air_Gate);
   14: XIC(Open_Treat_Air_Gate)TON(Bin.tmrStartDelay,10000,10000);
   15: [XIO(Open_Treat_Air_Gate) ,EQU(Treat_Batch_Status,8) ]TON(Bin.tmrStopDelay,5000,0);
   16: [XIC(Bin.tmrStartDelay.DN) ,XIC(Bin.tmrStopDelay.TT) ]OTE(Open_Treat_Air_Gate_Ready);
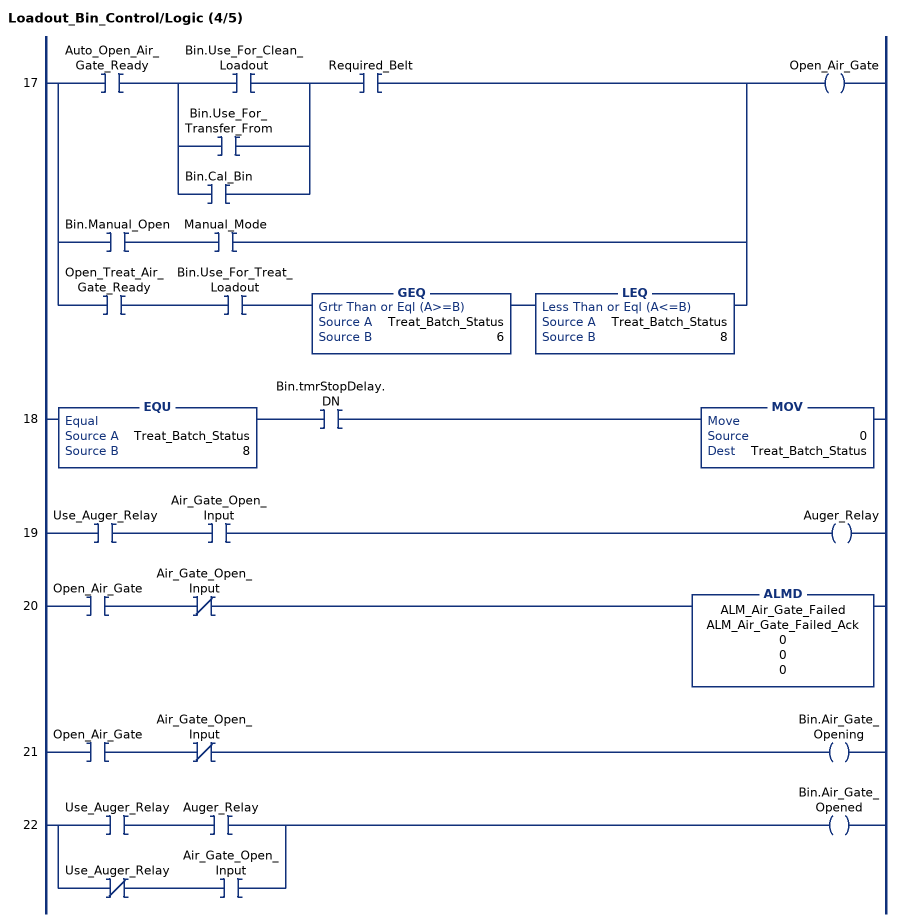
   17: [XIC(Auto_Open_Air_Gate_Ready) [XIC(Bin.Use_For_Clean_Loadout) ,XIC(Bin.Use_For_Transfer_From) ,XIC(Bin.Cal_Bin) ] XIC(Required_Belt) ,XIC(Bin.Manual_Open) XIC(Manual_Mode) ,XIC(Open_Treat_Air_Gate_Ready) XIC(Bin.Use_For_Treat_Loadout) GEQ(Treat_Batch_Status,6) LEQ(Treat_Batch_Status,8) ]OTE(Open_Air_Gate);
   18: EQU(Treat_Batch_Status,8)XIC(Bin.tmrStopDelay.DN)MOV(0,Treat_Batch_Status);
   19: XIC(Use_Auger_Relay)XIC(Air_Gate_Open_Input)OTE(Auger_Relay);
   20: XIC(Open_Air_Gate)XIO(Air_Gate_Open_Input)ALMD(ALM_Air_Gate_Failed,ALM_Air_Gate_Failed_Ack,0,0,0);
   21: XIC(Open_Air_Gate)XIO(Air_Gate_Open_Input)OTE(Bin.Air_Gate_Opening);
   22: [XIC(Use_Auger_Relay) XIC(Auger_Relay) ,XIO(Use_Auger_Relay) XIC(Air_Gate_Open_Input) ]OTE(Bin.Air_Gate_Opened);
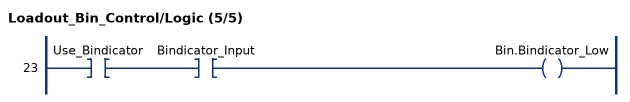
   23: XIC(Use_Bindicator)XIC(Bindicator_Input)OTE(Bin.Bindicator_Low);
END_ROUTINE
END_ADD_ON_INSTRUCTION
